FUNCTION_BLOCK Controle_Revezamento_3_HMI (* Service Interface Function Block Type *)
  (* Standard: 61499-2 *)
  (* Version 1.0, 21/10/2026, Hidryco, Hidryco, IHM do Controle_Revezamento_3 *)
  PACKAGE Hidryco.HidrycoLib;
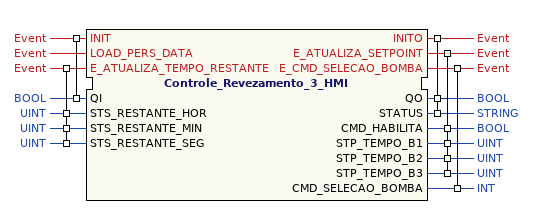
  EVENT_INPUT
    INIT WITH QI;
    LOAD_PERS_DATA; (* Reenvia os parametros persistentes *)
    E_ATUALIZA_TEMPO_RESTANTE WITH STS_RESTANTE_HOR, STS_RESTANTE_MIN, STS_RESTANTE_SEG; (* Status do processo *)
  END_EVENT
  EVENT_OUTPUT
    INITO WITH QO, STATUS;
    E_ATUALIZA_SETPOINT WITH CMD_HABILITA, STP_TEMPO_B1, STP_TEMPO_B2, STP_TEMPO_B3; (* Ajustes (IHM/OPC UA e LOAD_PERS_DATA) *)
    E_CMD_SELECAO_BOMBA WITH CMD_SELECAO_BOMBA; (* Ajustes (IHM/OPC UA e LOAD_PERS_DATA) *)
  END_EVENT
  VAR_INPUT
    QI : BOOL;
    STS_RESTANTE_HOR : UINT; (* Tempo para a troca da principal (h) *)
    STS_RESTANTE_MIN : UINT; (* Tempo para a troca da principal (min) *)
    STS_RESTANTE_SEG : UINT; (* Tempo para a troca da principal (s) *)
  END_VAR
  VAR_OUTPUT
    QO : BOOL; (* Event Output Qualifier *)
    STATUS : STRING; (* Service Status *)
    CMD_HABILITA : BOOL; (* Troca da principal por tempo *)
    STP_TEMPO_B1 : UINT; (* Horas do equipamento 1 como principal *)
    STP_TEMPO_B2 : UINT; (* Horas do equipamento 2 como principal *)
    STP_TEMPO_B3 : UINT; (* Horas do equipamento 3 como principal *)
    CMD_SELECAO_BOMBA : INT; (* Bomba principal *)
  END_VAR
  SERVICE /
    SEQUENCE 
    END_SEQUENCE
  END_SERVICE
END_FUNCTION_BLOCK
